RoboDK station: ur5e_station.rdk

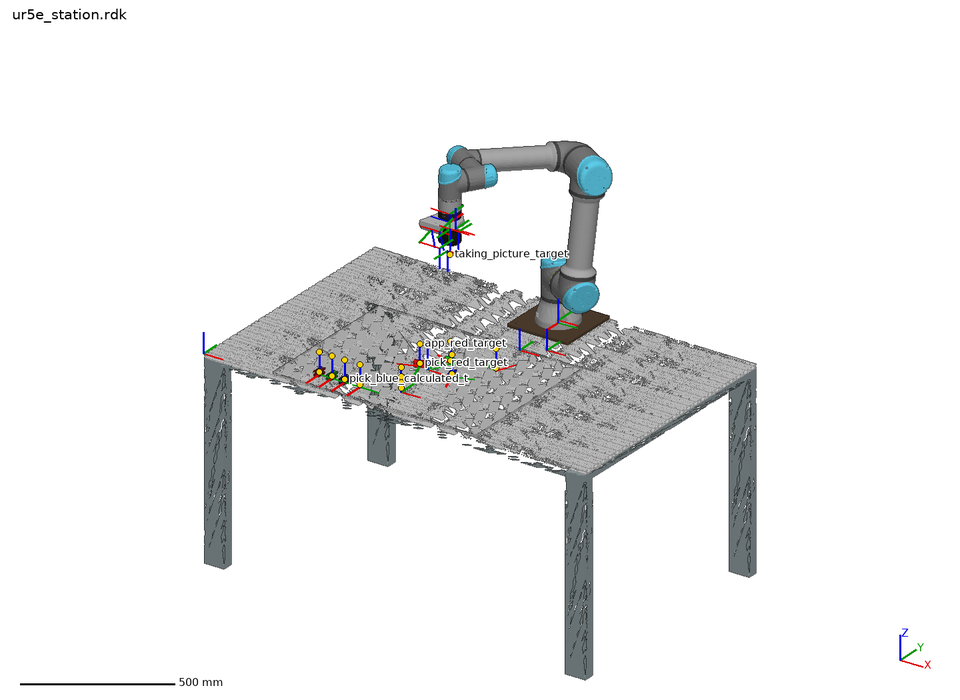
[picture v0: the station drawn from its stored meshes, robots at their saved joint values, targets as dots, program paths as lines]
Station ur5e_station (saved by RoboDK 5.6.7). Poses are relative to the parent item; angles as X-Y-Z fixed-axis rotations.
Station parameters (name, value as stored): PATH_MATLAB, C:\BRO_IRO_LAB\bro_iro_3_visionpnp-WS2024, IO_5, 1, IO_7, 1, RUN_MODE, 0, PATH_MATLAB_IMAGES, C:\BRO_IRO_LAB\bro_iro_3_visionpnp-WS2024\Images\, Palletizing Plugin
  - frame table_frame at (0, 1000, 0) mm
    - object table_object at (0, 0, 0) mm, size 1500 x 960.1 x 750 mm, geometry from Table.sld
    - frame white_frame at (670, 300, 10) mm
      - object white_object at (0, 0, 0) mm, size 800 x 600 x 10 mm, geometry from White Plate.STEP
    - frame robot_plate_frame at (806, 840, 0) mm, rotated rx 0 ry 0 rz -90 deg
      - object robot_plate_object at (0, 0, 0) mm, size 240 x 240 x 10 mm, 12 curves, geometry from 200731_v2_ur5e_bodenplatte_cad_jt.igs
    - frame UR5e Base at (806, 840, 10) mm
      - robot UR5e: 6 axes, payload 5 kg, reach 850 mm, repeatability 0.03 mm, weight 18.4 kg
          modified DH rows (alpha deg, a mm, theta deg, d mm): 0, 0, 0, 162.5; 90, 0, 180, 0; 0, 425, 0, 0; 0, 392.25, 0, 133.3; -90, 0, 0, 99.7; 90, 0, 180, 99.6
          joint limits [-360, -360, -360, -360, -360, -360] to [360, 360, 360, 360, 360, 360]; home [0, -90, -90, 0, 90, 0]; saved at [58.943, -96.374, 88.637, 277.653, -90, 148.979]
        - frame gripper_frame at (0, 0, 12) mm, rotated rx 0 ry 0 rz 180 deg
          - object Hand-E_IO_Coupling at (0, 0, -8) mm, size 75 x 105.3 x 17 mm, geometry from Hand-E_IO_Coupling.STEP
          - frame RobotiQ Hand-E Gripper Base at (0, 0, 0) mm
            - robot RobotiQ Hand-E Gripper: 1 axes
                joint limits [0] to [50]; home [0]; saved at [50]
          - frame Camera_and_Holder_Frame at (0, 0, 29) mm, rotated rx 90 ry 0 rz 90 deg
            - object hande_realsense_v5 at (0, 0, 0) mm, size 76.3 x 20 x 134.5 mm, geometry from hande_realsense_v5.stl
            - object counterpart holder v5 at (0, 0, 0) mm, size 42.7 x 20 x 99.3 mm, geometry from counterpart holder v5.stl
            - frame Intel RealSense D435 Frame at (-55.72, 12.9, 32.5) mm, rotated rx 0 ry 90 rz 75 deg
              - object Intel RealSense D435 at (0, 0, 0) mm, size 89.8 x 25 x 25.1 mm, geometry from Intel-RealSense-D435.sld
              - frame Camera Frame at (32.5, 0, 0) mm, rotated rx 0 ry 0 rz 180 deg
        - frame old___camera_frame_realsense at (0, -31, 77.7) mm, rotated rx -180 ry 0 rz 0 deg
          - object camera_holder_object at (0, 0, 0) mm, size 100 x 30 x 31 mm, geometry from Camera_holder.stl
          - frame Intel RealSense D435 Frame at (0, 17.5, -17) mm, rotated rx 180 ry 0 rz 180 deg
            - object Intel RealSense D435 at (0, 0, 0) mm, size 89.8 x 25 x 25.1 mm, geometry from Intel-RealSense-D435.sld
            - frame Camera Frame at (32.5, 0, 0) mm, rotated rx 0 ry 0 rz 180 deg
        - frame old___camera_frame_k4a at (0, 58, 111) mm, rotated rx 0 ry 0 rz 180 deg
          - object 2203___kamerahalterung at (0, 0, 0) mm, size 103 x 46.2 x 132 mm, geometry from 2203___kamerahalterung.step
          - frame camera_frame_k4a_rgb at (-32, 0, 0) mm, rotated rx 0 ry 0 rz 180 deg
            - camera 4ka_camera_rgb_768x432
        - tool gripper_tcp, TCP at (0, 0, 158.3) mm
        - tool camera_tcp_realsense_rgb, TCP at (0, 55.72, 53.9) mm, rotated rx -15 ry 0 rz 180 deg
        - tool camera_tcp_k4a_rgb, TCP at (32, 58, 111) mm
      - frame red_part_frame at (-170, -535, 0) mm, rotated rx 0 ry 0 rz -160 deg
        - target pick_red_target (Cartesian target) at (0, 0, 10) mm, rotated rx -180 ry 0 rz -90 deg; joints [57.289, -67.905, 115.158, 222.749, -89.903, 37.63] of UR5e
        - target app_red_target (Cartesian target) at (0, 0, 80) mm, rotated rx -180 ry 0 rz -90 deg; joints [57.298, -74.793, 111.478, 233.318, -89.861, 37.606] of UR5e
        - object red_object at (0, 0, 0) mm, size 40 x 20 x 20 mm, 1 curves, geometry from part.sld
      - frame green_part_frame at (-100, -460, 0) mm, rotated rx 0 ry 0 rz 160 deg
        - target pick_green_target (Cartesian target) at (0, 0, 10) mm, rotated rx -180 ry 0 rz -90 deg; joints [61.683, -75.138, 126.182, 218.958, -89.896, 81.259] of UR5e
        - target app_green_target (Cartesian target) at (0, 0, 80) mm, rotated rx -180 ry 0 rz -90 deg; joints [61.692, -83.219, 122.096, 231.124, -89.843, 81.229] of UR5e
        - object green_object at (0, 0, 0) mm, size 40 x 20 x 20 mm, 1 curves, geometry from part.sld
      - frame blue_part_frame at (-40, -540, 0) mm, rotated rx 0 ry 0 rz -70 deg
        - target pick_blue_target (Cartesian target) at (0, 0, 10) mm, rotated rx -180 ry 0 rz -90 deg; joints [71.724, -67.432, 114.399, 223.036, -89.903, -39.482] of UR5e
        - target app_blue_target (Cartesian target) at (0, 0, 80) mm, rotated rx 180 ry 0 rz -90 deg; joints [71.733, -74.25, 110.739, 233.514, -89.863, -39.505] of UR5e
        - object blue_object at (0, 0, 0) mm, size 40 x 20 x 20 mm, 1 curves, geometry from part.sld
      - frame black_part_frame at (50, -420, 0) mm, rotated rx 0 ry 0 rz 70 deg
        - target pick_blue_target (Cartesian target) at (0, 0, 10) mm, rotated rx -180 ry 0 rz -90 deg; joints [71.724, -67.432, 114.399, 223.036, -89.903, -39.482] of UR5e
        - target app_blue_target (Cartesian target) at (0, 0, 80) mm, rotated rx 180 ry 0 rz -90 deg; joints [71.733, -74.25, 110.739, 233.514, -89.863, -39.505] of UR5e
        - object black_object at (0, 0, 0) mm, size 40 x 20 x 20 mm, 1 curves, geometry from part.sld
      - frame red_part_calculated_frame at (-400, -770, 0) mm, rotated rx 0 ry 0 rz -90 deg
        - target app_red_calculated_target (Cartesian target) at (0, 0, 80) mm, rotated rx 180 ry 0 rz 90 deg; joints [53.645, -30.276, 35.937, 264.342, -89.93, 143.733] of UR5e
        - target pick_red_calculated_target (Cartesian target) at (0, 0, 10) mm, rotated rx 180 ry 0 rz 90 deg; joints [53.633, -27.741, 41.336, 256.407, -89.931, 143.75] of UR5e
        - object red_calculated_object at (0, 0, 0) mm, size 40 x 20 x 20 mm, 1 curves, geometry from part.sld
      - frame green_part_calculated_frame at (-350, -770, 0) mm, rotated rx 0 ry 0 rz -90 deg
        - target app_green_calculated_target (Cartesian target) at (0, 0, 80) mm, rotated rx -180 ry 0 rz 90 deg; joints [56.406, -34.841, 44.707, 260.138, -89.922, 146.525] of UR5e
        - target pick_green_calculated_target (Cartesian target) at (0, 0, 10) mm, rotated rx 180 ry 0 rz 90 deg; joints [56.396, -31.78, 49.317, 252.466, -89.928, 146.541] of UR5e
        - object green_calculated_object at (0, 0, 0) mm, size 40 x 20 x 20 mm, 1 curves, geometry from part.sld
      - frame blue_part_calculated_frame at (-300, -770, 0) mm, rotated rx 0 ry 0 rz -90 deg
        - target app_blue_calculated_target (Cartesian target) at (0, 0, 80) mm, rotated rx 180 ry 0 rz 90 deg; joints [59.337, -38.337, 51.301, 257.038, -89.917, 149.479] of UR5e
        - target pick_blue_calculated_target (Cartesian target) at (0, 0, 10) mm, rotated rx 180 ry 0 rz 90 deg; joints [59.327, -34.941, 55.503, 249.441, -89.925, 149.494] of UR5e
        - object blue_calculated_object at (0, 0, 0) mm, size 40 x 20 x 20 mm, 1 curves, geometry from part.sld
      - frame black_part_calculated_frame at (-240, -770, 0) mm, rotated rx 0 ry 0 rz -90 deg
        - target app_blue_calculated_target (Cartesian target) at (0, 0, 80) mm, rotated rx 180 ry 0 rz 90 deg; joints [59.337, -38.337, 51.301, 257.038, -89.917, 149.479] of UR5e
        - target pick_blue_calculated_target (Cartesian target) at (0, 0, 10) mm, rotated rx 180 ry 0 rz 90 deg; joints [59.327, -34.941, 55.503, 249.441, -89.925, 149.494] of UR5e
        - object black_calculated_object at (0, 0, 0) mm, size 40 x 20 x 20 mm, 1 curves, geometry from part.sld
      - frame place_frame at (-110, -725, 0.5) mm
        - target app_place_target (Cartesian target) at (0, 0, 90) mm, rotated rx 180 ry 0 rz 0 deg; joints [71.526, -48.414, 68.114, 250.303, -89.902, 161.72] of UR5e
        - target place_red_target (Cartesian target) at (0, 0, 15) mm, rotated rx 180 ry 0 rz 0 deg; joints [70.899, -47.844, 78.868, 238.976, -90, 160.899] of UR5e
        - target place_green_target (Cartesian target) at (0, 0, 35) mm, rotated rx 180 ry 0 rz 0 deg; joints [70.899, -49.216, 78.005, 241.211, -90, 160.899] of UR5e
        - target place_blue_target (Cartesian target) at (0, 0, 55) mm, rotated rx 180 ry 0 rz 0 deg; joints [70.899, -50.498, 76.999, 243.499, -90, 160.899] of UR5e
      - frame camara_calibration at (120, -236, 20) mm
        - frame Top_R at (-71, -50, 0) mm
          - object blue_object at (-20, -10, -20) mm, size 40 x 20 x 20 mm, 1 curves, geometry from part.sld
        - frame Top_L at (-349, -50, 0) mm
          - object blue_object at (20, -10, -20) mm, size 40 x 20 x 20 mm, 1 curves, geometry from part.sld
        - frame Bot_R at (-71, -247, 0) mm
          - object blue_object at (-20, 10, -20) mm, size 40 x 20 x 20 mm, 1 curves, geometry from part.sld
        - frame Bot_L at (-349, -247, 0) mm
          - object blue_object at (20, 10, -20) mm, size 40 x 20 x 20 mm, 1 curves, geometry from part.sld
      - target taking_picture_target (Cartesian target) at (-113.59, -447.06, 379.92) mm, rotated rx -179.93 ry -0.04 rz 179.96 deg; joints [58.759, -96.576, 90.28, 276.216, -89.784, -31.072] of UR5e
      - target taking_picture_target_k4a (Cartesian target) at (-113.61, -447.05, 379.92) mm, rotated rx 179.93 ry 0.04 rz -0.04 deg; joints [58.76, -96.41, 88.62, 277.71, -89.79, 148.92] of UR5e
    - frame gripper_move_frame at (0, 0, 0) mm
      - target open_gripper_full_target (joint target) at (692.39, 392.95, 386.22) mm, rotated rx -179.93 ry -0.04 rz 179.96 deg; joints [50, 11.333, 12.677, 10, 14.01, 14.333] of RobotiQ Hand-E Gripper
      - target open_gripper_20mm_target (Cartesian target) at (692.39, 392.95, 386.22) mm, rotated rx -179.93 ry -0.04 rz 179.96 deg; joints [20, 0, 0, 0, 0, 0] of RobotiQ Hand-E Gripper
      - target close_gripper_full_target (joint target) at (692.39, 392.95, 386.22) mm, rotated rx -179.93 ry -0.04 rz 179.96 deg; joints [0, 0, 0, 0, 0, 0] of RobotiQ Hand-E Gripper
  - folder program
    - folder robodk_code
      - folder pick_color_sim
        - program pick_red_sim (1 instructions, listed below)
        - program pick_green_sim (1 instructions, listed below)
        - program pick_blue_sim (1 instructions, listed below)
      - folder place_color_sim
        - program place_red_sim (1 instructions, listed below)
        - program place_blue_sim (1 instructions, listed below)
        - program place_green_sim (1 instructions, listed below)
      - folder gripper_programs
        - program HandE_CLOSE_SIM (1 instructions, listed below)
        - program HandE_OPEN_SIM (1 instructions, listed below)
        - program HandE_OPEN_SIM_20mm (1 instructions, listed below)
        - program HandE_OPEN_DIO (3 instructions, listed below)
        - program HandE_CLOSE_DIO (3 instructions, listed below)
        - program Hand-E_DO_ACTIVATE (9 instructions, listed below)
      - program UR5e_HOME_SIM (3 instructions, listed below)
      - program UR5e_HOME_REL (3 instructions, listed below)
    - folder python_code
      - Python program 4ka_sim (listed below)
      - Python program 4ka_real (listed below)
      - Python program realsense_sim (listed below)
      - Python program realsense_real_bkup (listed below)
      - Python program realsense_real (listed below)
      - Python program hande_open_gripper (listed below)
      - Python program hande_close_gripper (listed below)
      - Python program hande_activate_gripper (listed below)
    - program replace_all_objects (1 instructions, listed below)
    - program Main (7 instructions, listed below)
  - camera Camera 2
  - camera Kamera3
  - camera Kamera4
  - camera Kamera5
  - program open_gripper (1 instructions, listed below)
  - program close_gripper (2 instructions, listed below)
  - camera Camera 6

--- program pick_red_sim (robot UR5e) ---
  Attach to gripper_tcp

--- program pick_green_sim (robot UR5e) ---
  Attach to gripper_tcp

--- program pick_blue_sim (robot UR5e) ---
  Attach to gripper_tcp

--- program place_red_sim (robot UR5e) ---
  Detach from gripper_tcp

--- program place_blue_sim (robot UR5e) ---
  Detach from gripper_tcp

--- program place_green_sim (robot UR5e) ---
  Detach from gripper_tcp

--- program HandE_CLOSE_SIM (robot RobotiQ Hand-E Gripper) ---
  MoveJ (close_gripper_full_target)

--- program HandE_OPEN_SIM (robot RobotiQ Hand-E Gripper) ---
  MoveJ (open_gripper_full_target)

--- program HandE_OPEN_SIM_20mm (robot RobotiQ Hand-E Gripper) ---
  MoveJ (open_gripper_20mm_target)

--- program HandE_OPEN_DIO (robot UR5e) ---
  Call HandE_OPEN_SIM
  Set IO_6=1
  Pause 1.0 s

--- program HandE_CLOSE_DIO (robot UR5e) ---
  Call HandE_OPEN_SIM_20mm
  Set IO_6=0
  Pause 1.0 s

--- program Hand-E_DO_ACTIVATE (robot UR5e) ---
  Call HandE_CLOSE_SIM
  Set IO_6=1
  Pause 20 ms
  Set IO_6=0
  Pause 20 ms
  Set IO_7=1
  Pause 20 ms
  Set IO_7=0
  Pause 2.0 s

--- program UR5e_HOME_SIM (robot UR5e) ---
  Set Ref.: ur5e_frame -> UR5e Base
  Set Tool: gripper_tcp
  MoveJ (taking_picture_target_k4a)

--- program UR5e_HOME_REL (robot UR5e) ---
  Set Ref.: ur5e_frame -> UR5e Base
  Set Tool: gripper_tcp
  MoveJ (taking_picture_target_k4a)

--- Python program 4ka_sim ---
# This macro provokes taking a snapshot from a simulated 2D camera
#
from robolink import *    # API to communicate with RoboDK
from robodk import *      # basic matrix operations
RDK = Robolink()

#RDK.Cam2D_Close()

#camera = "r1s" #realsense
camera = "k4a" #Kinect

if camera == "r1s":
    camref = RDK.Item('camera_tcp_realsense_rgb',ITEM_TYPE_TOOL)
    cam_id = RDK.Cam2D_Add(camref, 'FOCAL_LENGHT=5 FOV=45 FAR_LENGHT=2000 SIZE=640x480')
elif camera == "k4a":
    camref = RDK.Item('camera_tcp_k4a_rgb',ITEM_TYPE_TOOL)
    cam_id = RDK.Cam2D_Add(camref, 'FOCAL_LENGHT=5 FOV=59 FAR_LENGHT=500 SIZE=768x432')

pause(1)

file_name = RDK.getParam('PATH_MATLAB_IMAGES') + "\Snap_sim.jpg"
RDK.Cam2D_Snapshot(file_name)
RDK.Cam2D_Close()

print("Saving camera snapshot to the file:" + file_name)

--- Python program 4ka_real ---
### Python 3 for the Azure-Kinect-Sensor-SDK
### https://github.com/etiennedub/pyk4a
### pip install pyk4a

### Other packages
### pip install numpy
### pip install opencv-python

import datetime
import numpy as np
import cv2
import pyk4a
#from pyk4a import Config, PyK4A

from robolink import *    # API to communicate with RoboDK
from robodk import *      # basic matrix operations
RDK = Robolink()
path = RDK.getParam('PATH_MATLAB')
print (path)
path = path + "\Images\\"
print (path)

def get_picture_azure(k4a):
    #### Position for taking Picture: MoveJ([71.03, -82.70, 82.13, 270.57, -89.82, -18.82]) #XYZRXRYRZ# -> -49.993, -550.003, 339.987, -0.002, 180.000, 0.002
    capture = k4a.get_capture()
    if np.any(capture.color):
        pic = capture.color[:,:,:3]
        #cv2.imshow("k4a", pic)
        #cv2.waitKey(0)
        pic = np.ascontiguousarray(pic)
    return pic


################

if __name__ == "__main__":
    #datetime object
    dt = datetime.datetime.now()
    print ("Start Time : "+ dt.strftime("%d_%m_%Y_%H_%M_%S"))

    k4a = pyk4a.PyK4A(
            pyk4a.Config(
                color_resolution=pyk4a.ColorResolution.RES_2160P,
                depth_mode=pyk4a.DepthMode.NFOV_UNBINNED,
                camera_fps= pyk4a.FPS.FPS_30,
                wired_sync_mode=pyk4a.WiredSyncMode.STANDALONE,
                synchronized_images_only=True,
        )
    )
    k4a.start()



    id = 0
    # print(k4a.calibration.get_camera_matrix(1))
    # print(k4a.calibration.get_distortion_coefficients(1))
    poses = []
    test=1
    while(test==1):
        #c = input("Press enter to take picture...")
        img = get_picture_azure(k4a)
        cv2.imshow("Camera taken",cv2.resize(img,(768,432)))
        #cv2.imwrite(path+str(id)+"_Image.png",img)
        cv2.imwrite(path+"Snap_real.png",cv2.resize(img,(768,432)))
        #cv2.waitKey(100)
        test=0




    dt = datetime.datetime.now()
    print ("Start Time : "+ dt.strftime("%d_%m_%Y_%H_%M_%S"))

--- Python program realsense_sim ---
# This macro provokes taking a snapshot from a simulated 2D camera
#
from robolink import *    # API to communicate with RoboDK
from robodk import *      # basic matrix operations
RDK = Robolink()

#RDK.Cam2D_Close()

camera = "r1s" #realsense
#camera = "k4a" #Kinect

if camera == "r1s":
    camref = RDK.Item('camera_tcp_realsense_rgb',ITEM_TYPE_TOOL)
    cam_id = RDK.Cam2D_Add(camref, 'FOCAL_LENGHT=5 FOV=45 FAR_LENGHT=2000 SIZE=640x480')
elif camera == "k4a":
    camref = RDK.Item('camera_tcp_k4a_rgb',ITEM_TYPE_TOOL)
    cam_id = RDK.Cam2D_Add(camref, 'FOCAL_LENGHT=5 FOV=59 FAR_LENGHT=500 SIZE=768x432')

pause(1)

file_name = RDK.getParam('PATH_MATLAB_IMAGES') + "/Snap_sim.jpg"
RDK.Cam2D_Snapshot(file_name)
RDK.Cam2D_Close()

print("Saving camera snapshot to the file:" + file_name)

--- Python program realsense_real_bkup ---
#import appropriate python modules to the program
import numpy as np
import cv2
from matplotlib import pyplot as plt
import pyrealsense2
from realsense_depth import *
import random

# initialization

# Initialize Camera Intel Realsense
dc = DepthCamera()




cv2.namedWindow("frame")
num = 0
rand = random.randint(0,50)


while True:

    ret, depth_frame, frame = dc.get_frame()

    k = cv2.waitKey(1) & 0xFF


    if k == ord('i'):

        path = "D:\FHWS\Student work\Competition\New Lab\Third submission\ur5e_vision_lab\Images\Snap_real.jpg"

        state = cv2.imwrite(path,frame)
        print state
        num = num + 1
    cv2.imshow("frame", frame)

    # break when user pressing ESC
    if k == 27:
        break

cv2.destroyAllWindows()

--- Python program realsense_real ---
#import appropriate python modules to the program
import numpy as np
import cv2
import pyrealsense2 as rs
import time

from robolink import *    # API to communicate with RoboDK
from robodk import *      # basic matrix operation

#path setup for image file
RDK = Robolink()
path = RDK.getParam('PATH_MATLAB')
print (path)
path = path + "\Images\\"
print (path)

try:
    #Intel Realsense Create a context object. This object owns the handles to all connected realsense devices
    pipeline = rs.pipeline()

    # Configure streams
    config = rs.config()

    # Get device product line for setting a supporting resolution
    pipeline_wrapper = rs.pipeline_wrapper(pipeline)
    pipeline_profile = config.resolve(pipeline_wrapper)
    device = pipeline_profile.get_device()
    device_product_line = str(device.get_info(rs.camera_info.product_line))

    found_rgb = False
    for s in device.sensors:
        if s.get_info(rs.camera_info.name) == 'RGB Camera':
            found_rgb = True
            break
    if not found_rgb:
        print("The demo requires Depth camera with Color sensor")
        exit(0)

    #set up streams
    #depth stream with fixed res : config.enable_stream(rs.stream.depth, 640, 480, rs.format.z16, 30)

    if device_product_line == 'L500':
        config.enable_stream(rs.stream.color, 960, 540, rs.format.bgr8, 30)
    else:
        config.enable_stream(rs.stream.color, 640, 480, rs.format.bgr8, 30)

    # Start streaming
    pipeline.start(config)

    time.sleep(3)

    # This call waits until a new coherent set of frames is available on a device
    # Calls to get_frame_data(...) and get_frame_timestamp(...) on a device will return stable values until wait_for_frames(...) is called
    frames = pipeline.wait_for_frames()
    print("pipeline created")
    color_frame = frames.get_color_frame()
    if not color_frame:
        print("failed to get frames")

    # Convert images to numpy arrays
    color_image = np.asanyarray(color_frame.get_data())

    # Show images
    cv2.namedWindow('RealSense', cv2.WINDOW_AUTOSIZE)
    cv2.imshow('RealSense', color_image)
    cv2.waitKey(1)

    #write image to file
    cv2.imwrite(path+"Snap_real.png",cv2.resize(color_image,(768,432)))


except Exception as e:
    print(e)
    pass

finally:
    # Stop streaming
    pipeline.stop()

--- Python program hande_open_gripper ---
"""Module to control Robotiq's grippers - tested with HAND-E"""

import socket
import threading
import time
from enum import Enum
from typing import Union, Tuple, OrderedDict

class RobotiqGripper:
    """
    Communicates with the gripper directly, via socket with string commands, leveraging string names for variables.
    """
    # WRITE VARIABLES (CAN ALSO READ)
    ACT = 'ACT'  # act : activate (1 while activated, can be reset to clear fault status)
    GTO = 'GTO'  # gto : go to (will perform go to with the actions set in pos, for, spe)
    ATR = 'ATR'  # atr : auto-release (emergency slow move)
    ADR = 'ADR'  # adr : auto-release direction (open(1) or close(0) during auto-release)
    FOR = 'FOR'  # for : force (0-255)
    SPE = 'SPE'  # spe : speed (0-255)
    POS = 'POS'  # pos : position (0-255), 0 = open
    # READ VARIABLES
    STA = 'STA'  # status (0 = is reset, 1 = activating, 3 = active)
    PRE = 'PRE'  # position request (echo of last commanded position)
    OBJ = 'OBJ'  # object detection (0 = moving, 1 = outer grip, 2 = inner grip, 3 = no object at rest)
    FLT = 'FLT'  # fault (0=ok, see manual for errors if not zero)

    ENCODING = 'UTF-8'  # ASCII and UTF-8 both seem to work

    class GripperStatus(Enum):
        """Gripper status reported by the gripper. The integer values have to match what the gripper sends."""
        RESET = 0
        ACTIVATING = 1
        # UNUSED = 2  # This value is currently not used by the gripper firmware
        ACTIVE = 3

    class ObjectStatus(Enum):
        """Object status reported by the gripper. The integer values have to match what the gripper sends."""
        MOVING = 0
        STOPPED_OUTER_OBJECT = 1
        STOPPED_INNER_OBJECT = 2
        AT_DEST = 3

    def __init__(self):
        """Constructor."""
        self.socket = None
        self.command_lock = threading.Lock()
        self._min_position = 0
        self._max_position = 255
        self._min_speed = 0
        self._max_speed = 255
        self._min_force = 0
        self._max_force = 255

    def connect(self, hostname: str, port: int, socket_timeout: float = 2.0) -> None:
        """Connects to a gripper at the given address.
        :param hostname: Hostname or ip.
        :param port: Port.
        :param socket_timeout: Timeout for blocking socket operations.
        """
        self.socket = socket.socket(socket.AF_INET, socket.SOCK_STREAM)
        self.socket.connect((hostname, port))
        self.socket.settimeout(socket_timeout)

    def disconnect(self) -> None:
        """Closes the connection with the gripper."""
        self.socket.close()

    def _set_vars(self, var_dict: OrderedDict[str, Union[int, float]]):
        """Sends the appropriate command via socket to set the value of n variables, and waits for its 'ack' response.
        :param var_dict: Dictionary of variables to set (variable_name, value).
        :return: True on successful reception of ack, false if no ack was received, indicating the set may not
        have been effective.
        """
        # construct unique command
        cmd = "SET"
        for variable, value in var_dict.items():
            cmd += f" {variable} {str(value)}"
        cmd += '\n'  # new line is required for the command to finish
        # atomic commands send/rcv
        with self.command_lock:
            self.socket.sendall(cmd.encode(self.ENCODING))
            data = self.socket.recv(1024)
        return self._is_ack(data)

    def _set_var(self, variable: str, value: Union[int, float]):
        """Sends the appropriate command via socket to set the value of a variable, and waits for its 'ack' response.
        :param variable: Variable to set.
        :param value: Value to set for the variable.
        :return: True on successful reception of ack, false if no ack was received, indicating the set may not
        have been effective.
        """
        return self._set_vars(OrderedDict([(variable, value)]))

    def _get_var(self, variable: str):
        """Sends the appropriate command to retrieve the value of a variable from the gripper, blocking until the
        response is received or the socket times out.
        :param variable: Name of the variable to retrieve.
        :return: Value of the variable as integer.
        """
        # atomic commands send/rcv
        with self.command_lock:
            cmd = f"GET {variable}\n"
            self.socket.sendall(cmd.encode(self.ENCODING))
            data = self.socket.recv(1024)

        # expect data of the form 'VAR x', where VAR is an echo of the variable name, and X the value
        # note some special variables (like FLT) may send 2 bytes, instead of an integer. We assume integer here
        var_name, value_str = data.decode(self.ENCODING).split()
        if var_name != variable:
            raise ValueError(f"Unexpected response {data} ({data.decode(self.ENCODING)}): does not match '{variable}'")
        value = int(value_str)
        return value

    @staticmethod
    def _is_ack(data: str):
        return data == b'ack'

    def _reset(self):
        """
        Reset the gripper.
        The following code is executed in the corresponding script function
        def rq_reset(gripper_socket="1"):
            rq_set_var("ACT", 0, gripper_socket)
            rq_set_var("ATR", 0, gripper_socket)

            while(not rq_get_var("ACT", 1, gripper_socket) == 0 or not rq_get_var("STA", 1, gripper_socket) == 0):
                rq_set_var("ACT", 0, gripper_socket)
                rq_set_var("ATR", 0, gripper_socket)
                sync()
            end

            sleep(0.5)
        end
        """
        self._set_var(self.ACT, 0)
        self._set_var(self.ATR, 0)
        while (not self._get_var(self.ACT) == 0 or not self._get_var(self.STA) == 0):
            self._set_var(self.ACT, 0)
            self._set_var(self.ATR, 0)
        time.sleep(0.5)


    def activate(self, auto_calibrate: bool = True):
        """Resets the activation flag in the gripper, and sets it back to one, clearing previous fault flags.
        :param auto_calibrate: Whether to calibrate the minimum and maximum positions based on actual motion.
        The following code is executed in the corresponding script function
        def rq_activate(gripper_socket="1"):
            if (not rq_is_gripper_activated(gripper_socket)):
                rq_reset(gripper_socket)

                while(not rq_get_var("ACT", 1, gripper_socket) == 0 or not rq_get_var("STA", 1, gripper_socket) == 0):
                    rq_reset(gripper_socket)
                    sync()
                end

                rq_set_var("ACT",1, gripper_socket)
            end
        end
        def rq_activate_and_wait(gripper_socket="1"):
            if (not rq_is_gripper_activated(gripper_socket)):
                rq_activate(gripper_socket)
                sleep(1.0)

                while(not rq_get_var("ACT", 1, gripper_socket) == 1 or not rq_get_var("STA", 1, gripper_socket) == 3):
                    sleep(0.1)
                end

                sleep(0.5)
            end
        end
        """
        if not self.is_active():
            self._reset()
            while (not self._get_var(self.ACT) == 0 or not self._get_var(self.STA) == 0):
                time.sleep(0.01)

            self._set_var(self.ACT, 1)
            time.sleep(1.0)
            while (not self._get_var(self.ACT) == 1 or not self._get_var(self.STA) == 3):
                time.sleep(0.01)

        # auto-calibrate position range if desired
        if auto_calibrate:
            self.auto_calibrate()

    def is_active(self):
        """Returns whether the gripper is active."""
        status = self._get_var(self.STA)
        return RobotiqGripper.GripperStatus(status) == RobotiqGripper.GripperStatus.ACTIVE

    def get_min_position(self) -> int:
        """Returns the minimum position the gripper can reach (open position)."""
        return self._min_position

    def get_max_position(self) -> int:
        """Returns the maximum position the gripper can reach (closed position)."""
        return self._max_position

    def get_open_position(self) -> int:
        """Returns what is considered the open position for gripper (minimum position value)."""
        return self.get_min_position()

    def get_closed_position(self) -> int:
        """Returns what is considered the closed position for gripper (maximum position value)."""
        return self.get_max_position()

    def is_open(self):
        """Returns whether the current position is considered as being fully open."""
        return self.get_current_position() <= self.get_open_position()

    def is_closed(self):
        """Returns whether the current position is considered as being fully closed."""
        return self.get_current_position() >= self.get_closed_position()

    def get_current_position(self) -> int:
        """Returns the current position as returned by the physical hardware."""
        return self._get_var(self.POS)

    def auto_calibrate(self, log: bool = True) -> None:
        """Attempts to calibrate the open and closed positions, by slowly closing and opening the gripper.
        :param log: Whether to print the results to log.
        """
        # first try to open in case we are holding an object
        (position, status) = self.move_and_wait_for_pos(self.get_open_position(), 64, 1)
        if RobotiqGripper.ObjectStatus(status) != RobotiqGripper.ObjectStatus.AT_DEST:
            raise RuntimeError(f"Calibration failed opening to start: {str(status)}")

        # try to close as far as possible, and record the number
        (position, status) = self.move_and_wait_for_pos(self.get_closed_position(), 64, 1)
        if RobotiqGripper.ObjectStatus(status) != RobotiqGripper.ObjectStatus.AT_DEST:
            raise RuntimeError(f"Calibration failed because of an object: {str(status)}")
        assert position <= self._max_position
        self._max_position = position

        # try to open as far as possible, and record the number
        (position, status) = self.move_and_wait_for_pos(self.get_open_position(), 64, 1)
        if RobotiqGripper.ObjectStatus(status) != RobotiqGripper.ObjectStatus.AT_DEST:
            raise RuntimeError(f"Calibration failed because of an object: {str(status)}")
        assert position >= self._min_position
        self._min_position = position

        if log:
            print(f"Gripper auto-calibrated to [{self.get_min_position()}, {self.get_max_position()}]")

    def move(self, position: int, speed: int, force: int) -> Tuple[bool, int]:
        """Sends commands to start moving towards the given position, with the specified speed and force.
        :param position: Position to move to [min_position, max_position]
        :param speed: Speed to move at [min_speed, max_speed]
        :param force: Force to use [min_force, max_force]
        :return: A tuple with a bool indicating whether the action it was successfully sent, and an integer with
        the actual position that was requested, after being adjusted to the min/max calibrated range.
        """

        def clip_val(min_val, val, max_val):
            return max(min_val, min(val, max_val))

        clip_pos = clip_val(self._min_position, position, self._max_position)
        clip_spe = clip_val(self._min_speed, speed, self._max_speed)
        clip_for = clip_val(self._min_force, force, self._max_force)

        # moves to the given position with the given speed and force
        var_dict = OrderedDict([(self.POS, clip_pos), (self.SPE, clip_spe), (self.FOR, clip_for), (self.GTO, 1)])
        return self._set_vars(var_dict), clip_pos

    def move_and_wait_for_pos(self, position: int, speed: int, force: int) -> Tuple[int, ObjectStatus]:  # noqa
        """Sends commands to start moving towards the given position, with the specified speed and force, and
        then waits for the move to complete.
        :param position: Position to move to [min_position, max_position]
        :param speed: Speed to move at [min_speed, max_speed]
        :param force: Force to use [min_force, max_force]
        :return: A tuple with an integer representing the last position returned by the gripper after it notified
        that the move had completed, a status indicating how the move ended (see ObjectStatus enum for details). Note
        that it is possible that the position was not reached, if an object was detected during motion.
        """
        set_ok, cmd_pos = self.move(position, speed, force)
        if not set_ok:
            raise RuntimeError("Failed to set variables for move.")

        # wait until the gripper acknowledges that it will try to go to the requested position
        while self._get_var(self.PRE) != cmd_pos:
            time.sleep(0.001)

        # wait until not moving
        cur_obj = self._get_var(self.OBJ)
        while RobotiqGripper.ObjectStatus(cur_obj) == RobotiqGripper.ObjectStatus.MOVING:
            cur_obj = self._get_var(self.OBJ)

        # report the actual position and the object status
        final_pos = self._get_var(self.POS)
        final_obj = cur_obj
        return final_pos, RobotiqGripper.ObjectStatus(final_obj)


if __name__ == '__main__':
    ip = "172.31.1.200"
    gripper = RobotiqGripper()
    print("Connecting to gripper...")
    gripper.connect(ip, 63352)
    #print("Activating gripper...")
    #gripper.activate()
    print("Open gripper...")
    gripper.move_and_wait_for_pos(0, 255, 255)

--- Python program hande_close_gripper ---
"""Module to control Robotiq's grippers - tested with HAND-E"""

import socket
import threading
import time
from enum import Enum
from typing import Union, Tuple, OrderedDict

class RobotiqGripper:
    """
    Communicates with the gripper directly, via socket with string commands, leveraging string names for variables.
    """
    # WRITE VARIABLES (CAN ALSO READ)
    ACT = 'ACT'  # act : activate (1 while activated, can be reset to clear fault status)
    GTO = 'GTO'  # gto : go to (will perform go to with the actions set in pos, for, spe)
    ATR = 'ATR'  # atr : auto-release (emergency slow move)
    ADR = 'ADR'  # adr : auto-release direction (open(1) or close(0) during auto-release)
    FOR = 'FOR'  # for : force (0-255)
    SPE = 'SPE'  # spe : speed (0-255)
    POS = 'POS'  # pos : position (0-255), 0 = open
    # READ VARIABLES
    STA = 'STA'  # status (0 = is reset, 1 = activating, 3 = active)
    PRE = 'PRE'  # position request (echo of last commanded position)
    OBJ = 'OBJ'  # object detection (0 = moving, 1 = outer grip, 2 = inner grip, 3 = no object at rest)
    FLT = 'FLT'  # fault (0=ok, see manual for errors if not zero)

    ENCODING = 'UTF-8'  # ASCII and UTF-8 both seem to work

    class GripperStatus(Enum):
        """Gripper status reported by the gripper. The integer values have to match what the gripper sends."""
        RESET = 0
        ACTIVATING = 1
        # UNUSED = 2  # This value is currently not used by the gripper firmware
        ACTIVE = 3

    class ObjectStatus(Enum):
        """Object status reported by the gripper. The integer values have to match what the gripper sends."""
        MOVING = 0
        STOPPED_OUTER_OBJECT = 1
        STOPPED_INNER_OBJECT = 2
        AT_DEST = 3

    def __init__(self):
        """Constructor."""
        self.socket = None
        self.command_lock = threading.Lock()
        self._min_position = 0
        self._max_position = 255
        self._min_speed = 0
        self._max_speed = 255
        self._min_force = 0
        self._max_force = 255

    def connect(self, hostname: str, port: int, socket_timeout: float = 2.0) -> None:
        """Connects to a gripper at the given address.
        :param hostname: Hostname or ip.
        :param port: Port.
        :param socket_timeout: Timeout for blocking socket operations.
        """
        self.socket = socket.socket(socket.AF_INET, socket.SOCK_STREAM)
        self.socket.connect((hostname, port))
        self.socket.settimeout(socket_timeout)

    def disconnect(self) -> None:
        """Closes the connection with the gripper."""
        self.socket.close()

    def _set_vars(self, var_dict: OrderedDict[str, Union[int, float]]):
        """Sends the appropriate command via socket to set the value of n variables, and waits for its 'ack' response.
        :param var_dict: Dictionary of variables to set (variable_name, value).
        :return: True on successful reception of ack, false if no ack was received, indicating the set may not
        have been effective.
        """
        # construct unique command
        cmd = "SET"
        for variable, value in var_dict.items():
            cmd += f" {variable} {str(value)}"
        cmd += '\n'  # new line is required for the command to finish
        # atomic commands send/rcv
        with self.command_lock:
            self.socket.sendall(cmd.encode(self.ENCODING))
            data = self.socket.recv(1024)
        return self._is_ack(data)

    def _set_var(self, variable: str, value: Union[int, float]):
        """Sends the appropriate command via socket to set the value of a variable, and waits for its 'ack' response.
        :param variable: Variable to set.
        :param value: Value to set for the variable.
        :return: True on successful reception of ack, false if no ack was received, indicating the set may not
        have been effective.
        """
        return self._set_vars(OrderedDict([(variable, value)]))

    def _get_var(self, variable: str):
        """Sends the appropriate command to retrieve the value of a variable from the gripper, blocking until the
        response is received or the socket times out.
        :param variable: Name of the variable to retrieve.
        :return: Value of the variable as integer.
        """
        # atomic commands send/rcv
        with self.command_lock:
            cmd = f"GET {variable}\n"
            self.socket.sendall(cmd.encode(self.ENCODING))
            data = self.socket.recv(1024)

        # expect data of the form 'VAR x', where VAR is an echo of the variable name, and X the value
        # note some special variables (like FLT) may send 2 bytes, instead of an integer. We assume integer here
        var_name, value_str = data.decode(self.ENCODING).split()
        if var_name != variable:
            raise ValueError(f"Unexpected response {data} ({data.decode(self.ENCODING)}): does not match '{variable}'")
        value = int(value_str)
        return value

    @staticmethod
    def _is_ack(data: str):
        return data == b'ack'

    def _reset(self):
        """
        Reset the gripper.
        The following code is executed in the corresponding script function
        def rq_reset(gripper_socket="1"):
            rq_set_var("ACT", 0, gripper_socket)
            rq_set_var("ATR", 0, gripper_socket)

            while(not rq_get_var("ACT", 1, gripper_socket) == 0 or not rq_get_var("STA", 1, gripper_socket) == 0):
                rq_set_var("ACT", 0, gripper_socket)
                rq_set_var("ATR", 0, gripper_socket)
                sync()
            end

            sleep(0.5)
        end
        """
        self._set_var(self.ACT, 0)
        self._set_var(self.ATR, 0)
        while (not self._get_var(self.ACT) == 0 or not self._get_var(self.STA) == 0):
            self._set_var(self.ACT, 0)
            self._set_var(self.ATR, 0)
        time.sleep(0.5)


    def activate(self, auto_calibrate: bool = True):
        """Resets the activation flag in the gripper, and sets it back to one, clearing previous fault flags.
        :param auto_calibrate: Whether to calibrate the minimum and maximum positions based on actual motion.
        The following code is executed in the corresponding script function
        def rq_activate(gripper_socket="1"):
            if (not rq_is_gripper_activated(gripper_socket)):
                rq_reset(gripper_socket)

                while(not rq_get_var("ACT", 1, gripper_socket) == 0 or not rq_get_var("STA", 1, gripper_socket) == 0):
                    rq_reset(gripper_socket)
                    sync()
                end

                rq_set_var("ACT",1, gripper_socket)
            end
        end
        def rq_activate_and_wait(gripper_socket="1"):
            if (not rq_is_gripper_activated(gripper_socket)):
                rq_activate(gripper_socket)
                sleep(1.0)

                while(not rq_get_var("ACT", 1, gripper_socket) == 1 or not rq_get_var("STA", 1, gripper_socket) == 3):
                    sleep(0.1)
                end

                sleep(0.5)
            end
        end
        """
        if not self.is_active():
            self._reset()
            while (not self._get_var(self.ACT) == 0 or not self._get_var(self.STA) == 0):
                time.sleep(0.01)

            self._set_var(self.ACT, 1)
            time.sleep(1.0)
            while (not self._get_var(self.ACT) == 1 or not self._get_var(self.STA) == 3):
                time.sleep(0.01)

        # auto-calibrate position range if desired
        if auto_calibrate:
            self.auto_calibrate()

    def is_active(self):
        """Returns whether the gripper is active."""
        status = self._get_var(self.STA)
        return RobotiqGripper.GripperStatus(status) == RobotiqGripper.GripperStatus.ACTIVE

    def get_min_position(self) -> int:
        """Returns the minimum position the gripper can reach (open position)."""
        return self._min_position

    def get_max_position(self) -> int:
        """Returns the maximum position the gripper can reach (closed position)."""
        return self._max_position

    def get_open_position(self) -> int:
        """Returns what is considered the open position for gripper (minimum position value)."""
        return self.get_min_position()

    def get_closed_position(self) -> int:
        """Returns what is considered the closed position for gripper (maximum position value)."""
        return self.get_max_position()

    def is_open(self):
        """Returns whether the current position is considered as being fully open."""
        return self.get_current_position() <= self.get_open_position()

    def is_closed(self):
        """Returns whether the current position is considered as being fully closed."""
        return self.get_current_position() >= self.get_closed_position()

    def get_current_position(self) -> int:
        """Returns the current position as returned by the physical hardware."""
        return self._get_var(self.POS)

    def auto_calibrate(self, log: bool = True) -> None:
        """Attempts to calibrate the open and closed positions, by slowly closing and opening the gripper.
        :param log: Whether to print the results to log.
        """
        # first try to open in case we are holding an object
        (position, status) = self.move_and_wait_for_pos(self.get_open_position(), 64, 1)
        if RobotiqGripper.ObjectStatus(status) != RobotiqGripper.ObjectStatus.AT_DEST:
            raise RuntimeError(f"Calibration failed opening to start: {str(status)}")

        # try to close as far as possible, and record the number
        (position, status) = self.move_and_wait_for_pos(self.get_closed_position(), 64, 1)
        if RobotiqGripper.ObjectStatus(status) != RobotiqGripper.ObjectStatus.AT_DEST:
            raise RuntimeError(f"Calibration failed because of an object: {str(status)}")
        assert position <= self._max_position
        self._max_position = position

        # try to open as far as possible, and record the number
        (position, status) = self.move_and_wait_for_pos(self.get_open_position(), 64, 1)
        if RobotiqGripper.ObjectStatus(status) != RobotiqGripper.ObjectStatus.AT_DEST:
            raise RuntimeError(f"Calibration failed because of an object: {str(status)}")
        assert position >= self._min_position
        self._min_position = position

        if log:
            print(f"Gripper auto-calibrated to [{self.get_min_position()}, {self.get_max_position()}]")

    def move(self, position: int, speed: int, force: int) -> Tuple[bool, int]:
        """Sends commands to start moving towards the given position, with the specified speed and force.
        :param position: Position to move to [min_position, max_position]
        :param speed: Speed to move at [min_speed, max_speed]
        :param force: Force to use [min_force, max_force]
        :return: A tuple with a bool indicating whether the action it was successfully sent, and an integer with
        the actual position that was requested, after being adjusted to the min/max calibrated range.
        """

        def clip_val(min_val, val, max_val):
            return max(min_val, min(val, max_val))

        clip_pos = clip_val(self._min_position, position, self._max_position)
        clip_spe = clip_val(self._min_speed, speed, self._max_speed)
        clip_for = clip_val(self._min_force, force, self._max_force)

        # moves to the given position with the given speed and force
        var_dict = OrderedDict([(self.POS, clip_pos), (self.SPE, clip_spe), (self.FOR, clip_for), (self.GTO, 1)])
        return self._set_vars(var_dict), clip_pos

    def move_and_wait_for_pos(self, position: int, speed: int, force: int) -> Tuple[int, ObjectStatus]:  # noqa
        """Sends commands to start moving towards the given position, with the specified speed and force, and
        then waits for the move to complete.
        :param position: Position to move to [min_position, max_position]
        :param speed: Speed to move at [min_speed, max_speed]
        :param force: Force to use [min_force, max_force]
        :return: A tuple with an integer representing the last position returned by the gripper after it notified
        that the move had completed, a status indicating how the move ended (see ObjectStatus enum for details). Note
        that it is possible that the position was not reached, if an object was detected during motion.
        """
        set_ok, cmd_pos = self.move(position, speed, force)
        if not set_ok:
            raise RuntimeError("Failed to set variables for move.")

        # wait until the gripper acknowledges that it will try to go to the requested position
        while self._get_var(self.PRE) != cmd_pos:
            time.sleep(0.001)

        # wait until not moving
        cur_obj = self._get_var(self.OBJ)
        while RobotiqGripper.ObjectStatus(cur_obj) == RobotiqGripper.ObjectStatus.MOVING:
            cur_obj = self._get_var(self.OBJ)

        # report the actual position and the object status
        final_pos = self._get_var(self.POS)
        final_obj = cur_obj
        return final_pos, RobotiqGripper.ObjectStatus(final_obj)


if __name__ == '__main__':
    ip = "172.31.1.200"
    gripper = RobotiqGripper()
    print("Connecting to gripper...")
    gripper.connect(ip, 63352)
    #print("Activating gripper...")
    #gripper.activate()
    print("Close gripper...")
    gripper.move_and_wait_for_pos(255, 255, 255)

--- Python program hande_activate_gripper ---
"""Module to control Robotiq's grippers - tested with HAND-E"""

import socket
import threading
import time
from enum import Enum
from typing import Union, Tuple, OrderedDict

class RobotiqGripper:
    """
    Communicates with the gripper directly, via socket with string commands, leveraging string names for variables.
    """
    # WRITE VARIABLES (CAN ALSO READ)
    ACT = 'ACT'  # act : activate (1 while activated, can be reset to clear fault status)
    GTO = 'GTO'  # gto : go to (will perform go to with the actions set in pos, for, spe)
    ATR = 'ATR'  # atr : auto-release (emergency slow move)
    ADR = 'ADR'  # adr : auto-release direction (open(1) or close(0) during auto-release)
    FOR = 'FOR'  # for : force (0-255)
    SPE = 'SPE'  # spe : speed (0-255)
    POS = 'POS'  # pos : position (0-255), 0 = open
    # READ VARIABLES
    STA = 'STA'  # status (0 = is reset, 1 = activating, 3 = active)
    PRE = 'PRE'  # position request (echo of last commanded position)
    OBJ = 'OBJ'  # object detection (0 = moving, 1 = outer grip, 2 = inner grip, 3 = no object at rest)
    FLT = 'FLT'  # fault (0=ok, see manual for errors if not zero)

    ENCODING = 'UTF-8'  # ASCII and UTF-8 both seem to work

    class GripperStatus(Enum):
        """Gripper status reported by the gripper. The integer values have to match what the gripper sends."""
        RESET = 0
        ACTIVATING = 1
        # UNUSED = 2  # This value is currently not used by the gripper firmware
        ACTIVE = 3

    class ObjectStatus(Enum):
        """Object status reported by the gripper. The integer values have to match what the gripper sends."""
        MOVING = 0
        STOPPED_OUTER_OBJECT = 1
        STOPPED_INNER_OBJECT = 2
        AT_DEST = 3

    def __init__(self):
        """Constructor."""
        self.socket = None
        self.command_lock = threading.Lock()
        self._min_position = 0
        self._max_position = 255
        self._min_speed = 0
        self._max_speed = 255
        self._min_force = 0
        self._max_force = 255

    def connect(self, hostname: str, port: int, socket_timeout: float = 2.0) -> None:
        """Connects to a gripper at the given address.
        :param hostname: Hostname or ip.
        :param port: Port.
        :param socket_timeout: Timeout for blocking socket operations.
        """
        self.socket = socket.socket(socket.AF_INET, socket.SOCK_STREAM)
        self.socket.connect((hostname, port))
        self.socket.settimeout(socket_timeout)

    def disconnect(self) -> None:
        """Closes the connection with the gripper."""
        self.socket.close()

    def _set_vars(self, var_dict: OrderedDict[str, Union[int, float]]):
        """Sends the appropriate command via socket to set the value of n variables, and waits for its 'ack' response.
        :param var_dict: Dictionary of variables to set (variable_name, value).
        :return: True on successful reception of ack, false if no ack was received, indicating the set may not
        have been effective.
        """
        # construct unique command
        cmd = "SET"
        for variable, value in var_dict.items():
            cmd += f" {variable} {str(value)}"
        cmd += '\n'  # new line is required for the command to finish
        # atomic commands send/rcv
        with self.command_lock:
            self.socket.sendall(cmd.encode(self.ENCODING))
            data = self.socket.recv(1024)
        return self._is_ack(data)

    def _set_var(self, variable: str, value: Union[int, float]):
        """Sends the appropriate command via socket to set the value of a variable, and waits for its 'ack' response.
        :param variable: Variable to set.
        :param value: Value to set for the variable.
        :return: True on successful reception of ack, false if no ack was received, indicating the set may not
        have been effective.
        """
        return self._set_vars(OrderedDict([(variable, value)]))

    def _get_var(self, variable: str):
        """Sends the appropriate command to retrieve the value of a variable from the gripper, blocking until the
        response is received or the socket times out.
        :param variable: Name of the variable to retrieve.
        :return: Value of the variable as integer.
        """
        # atomic commands send/rcv
        with self.command_lock:
            cmd = f"GET {variable}\n"
            self.socket.sendall(cmd.encode(self.ENCODING))
            data = self.socket.recv(1024)

        # expect data of the form 'VAR x', where VAR is an echo of the variable name, and X the value
        # note some special variables (like FLT) may send 2 bytes, instead of an integer. We assume integer here
        var_name, value_str = data.decode(self.ENCODING).split()
        if var_name != variable:
            raise ValueError(f"Unexpected response {data} ({data.decode(self.ENCODING)}): does not match '{variable}'")
        value = int(value_str)
        return value

    @staticmethod
    def _is_ack(data: str):
        return data == b'ack'

    def _reset(self):
        """
        Reset the gripper.
        The following code is executed in the corresponding script function
        def rq_reset(gripper_socket="1"):
            rq_set_var("ACT", 0, gripper_socket)
            rq_set_var("ATR", 0, gripper_socket)

            while(not rq_get_var("ACT", 1, gripper_socket) == 0 or not rq_get_var("STA", 1, gripper_socket) == 0):
                rq_set_var("ACT", 0, gripper_socket)
                rq_set_var("ATR", 0, gripper_socket)
                sync()
            end

            sleep(0.5)
        end
        """
        self._set_var(self.ACT, 0)
        self._set_var(self.ATR, 0)
        while (not self._get_var(self.ACT) == 0 or not self._get_var(self.STA) == 0):
            self._set_var(self.ACT, 0)
            self._set_var(self.ATR, 0)
        time.sleep(0.5)


    def activate(self, auto_calibrate: bool = True):
        """Resets the activation flag in the gripper, and sets it back to one, clearing previous fault flags.
        :param auto_calibrate: Whether to calibrate the minimum and maximum positions based on actual motion.
        The following code is executed in the corresponding script function
        def rq_activate(gripper_socket="1"):
            if (not rq_is_gripper_activated(gripper_socket)):
                rq_reset(gripper_socket)

                while(not rq_get_var("ACT", 1, gripper_socket) == 0 or not rq_get_var("STA", 1, gripper_socket) == 0):
                    rq_reset(gripper_socket)
                    sync()
                end

                rq_set_var("ACT",1, gripper_socket)
            end
        end
        def rq_activate_and_wait(gripper_socket="1"):
            if (not rq_is_gripper_activated(gripper_socket)):
                rq_activate(gripper_socket)
                sleep(1.0)

                while(not rq_get_var("ACT", 1, gripper_socket) == 1 or not rq_get_var("STA", 1, gripper_socket) == 3):
                    sleep(0.1)
                end

                sleep(0.5)
            end
        end
        """
        if not self.is_active():
            self._reset()
            while (not self._get_var(self.ACT) == 0 or not self._get_var(self.STA) == 0):
                time.sleep(0.01)

            self._set_var(self.ACT, 1)
            time.sleep(1.0)
            while (not self._get_var(self.ACT) == 1 or not self._get_var(self.STA) == 3):
                time.sleep(0.01)

        # auto-calibrate position range if desired
        if auto_calibrate:
            self.auto_calibrate()

    def is_active(self):
        """Returns whether the gripper is active."""
        status = self._get_var(self.STA)
        return RobotiqGripper.GripperStatus(status) == RobotiqGripper.GripperStatus.ACTIVE

    def get_min_position(self) -> int:
        """Returns the minimum position the gripper can reach (open position)."""
        return self._min_position

    def get_max_position(self) -> int:
        """Returns the maximum position the gripper can reach (closed position)."""
        return self._max_position

    def get_open_position(self) -> int:
        """Returns what is considered the open position for gripper (minimum position value)."""
        return self.get_min_position()

    def get_closed_position(self) -> int:
        """Returns what is considered the closed position for gripper (maximum position value)."""
        return self.get_max_position()

    def is_open(self):
        """Returns whether the current position is considered as being fully open."""
        return self.get_current_position() <= self.get_open_position()

    def is_closed(self):
        """Returns whether the current position is considered as being fully closed."""
        return self.get_current_position() >= self.get_closed_position()

    def get_current_position(self) -> int:
        """Returns the current position as returned by the physical hardware."""
        return self._get_var(self.POS)

    def auto_calibrate(self, log: bool = True) -> None:
        """Attempts to calibrate the open and closed positions, by slowly closing and opening the gripper.
        :param log: Whether to print the results to log.
        """
        # first try to open in case we are holding an object
        (position, status) = self.move_and_wait_for_pos(self.get_open_position(), 64, 1)
        if RobotiqGripper.ObjectStatus(status) != RobotiqGripper.ObjectStatus.AT_DEST:
            raise RuntimeError(f"Calibration failed opening to start: {str(status)}")

        # try to close as far as possible, and record the number
        (position, status) = self.move_and_wait_for_pos(self.get_closed_position(), 64, 1)
        if RobotiqGripper.ObjectStatus(status) != RobotiqGripper.ObjectStatus.AT_DEST:
            raise RuntimeError(f"Calibration failed because of an object: {str(status)}")
        assert position <= self._max_position
        self._max_position = position

        # try to open as far as possible, and record the number
        (position, status) = self.move_and_wait_for_pos(self.get_open_position(), 64, 1)
        if RobotiqGripper.ObjectStatus(status) != RobotiqGripper.ObjectStatus.AT_DEST:
            raise RuntimeError(f"Calibration failed because of an object: {str(status)}")
        assert position >= self._min_position
        self._min_position = position

        if log:
            print(f"Gripper auto-calibrated to [{self.get_min_position()}, {self.get_max_position()}]")

    def move(self, position: int, speed: int, force: int) -> Tuple[bool, int]:
        """Sends commands to start moving towards the given position, with the specified speed and force.
        :param position: Position to move to [min_position, max_position]
        :param speed: Speed to move at [min_speed, max_speed]
        :param force: Force to use [min_force, max_force]
        :return: A tuple with a bool indicating whether the action it was successfully sent, and an integer with
        the actual position that was requested, after being adjusted to the min/max calibrated range.
        """

        def clip_val(min_val, val, max_val):
            return max(min_val, min(val, max_val))

        clip_pos = clip_val(self._min_position, position, self._max_position)
        clip_spe = clip_val(self._min_speed, speed, self._max_speed)
        clip_for = clip_val(self._min_force, force, self._max_force)

        # moves to the given position with the given speed and force
        var_dict = OrderedDict([(self.POS, clip_pos), (self.SPE, clip_spe), (self.FOR, clip_for), (self.GTO, 1)])
        return self._set_vars(var_dict), clip_pos

    def move_and_wait_for_pos(self, position: int, speed: int, force: int) -> Tuple[int, ObjectStatus]:  # noqa
        """Sends commands to start moving towards the given position, with the specified speed and force, and
        then waits for the move to complete.
        :param position: Position to move to [min_position, max_position]
        :param speed: Speed to move at [min_speed, max_speed]
        :param force: Force to use [min_force, max_force]
        :return: A tuple with an integer representing the last position returned by the gripper after it notified
        that the move had completed, a status indicating how the move ended (see ObjectStatus enum for details). Note
        that it is possible that the position was not reached, if an object was detected during motion.
        """
        set_ok, cmd_pos = self.move(position, speed, force)
        if not set_ok:
            raise RuntimeError("Failed to set variables for move.")

        # wait until the gripper acknowledges that it will try to go to the requested position
        while self._get_var(self.PRE) != cmd_pos:
            time.sleep(0.001)

        # wait until not moving
        cur_obj = self._get_var(self.OBJ)
        while RobotiqGripper.ObjectStatus(cur_obj) == RobotiqGripper.ObjectStatus.MOVING:
            cur_obj = self._get_var(self.OBJ)

        # report the actual position and the object status
        final_pos = self._get_var(self.POS)
        final_obj = cur_obj
        return final_pos, RobotiqGripper.ObjectStatus(final_obj)


if __name__ == '__main__':
    ip = "172.31.1.200"
    gripper = RobotiqGripper()
    print("Connecting to gripper...")
    gripper.connect(ip, 63352)
    print("Activating gripper...")
    gripper.activate()
    #print("Close gripper...")
    #gripper.move_and_wait_for_pos(255, 255, 255)

--- program replace_all_objects (robot UR5e) ---
  Replace objects

--- program Main (robot UR5e) ---
  Call open_gripper_full
  Call pick_red
  Call place_red
  Call pick_green
  Call place_green
  Call pick_blue
  Call place_blue

--- program open_gripper (robot UR5e) ---
  Call rq_move_and_wait(255)

--- program close_gripper (robot UR5e) ---
  Call rq_move_and_wait( 0 )
  Pause 1.0 s
